FUNCTION_BLOCK DRIVE
  VAR_INPUT
    A : BOOL;
    B : BOOL;
    C : BOOL;
  END_VAR
  VAR_OUTPUT
    Y : BOOL;
  END_VAR

BEGIN
Y := A AND B AND C;
  //#ASSERT NOT Y OR (A AND B AND C) : P1
END_FUNCTION_BLOCK
